// TIA Portal V21 export
// export: Created 2026-11-10T07:26:50.592199Z, ExportSetting WithDefaults, DisplayName Totally Integrated Automation Portal, DisplayVersion V21 Update 3, DisplayName STEP 7 Professional, DisplayVersion V21 Update 3, DisplayName STEP 7 Safety, DisplayVersion V21, DisplayName Tech WebApplication, DisplayVersion V21, DisplayName WinCC Basic/Comfort/Advanced, DisplayVersion V21 Update 3, DisplayName WinCC Unified, DisplayVersion V21 Update 3
FUNCTION_BLOCK "FB_LadOperands"   // FB5, LAD
{ S7_Optimized_Access := 'TRUE' }
VERSION : 0.1
// stored: AutoNumber true, IsIECCheckEnabled false, IsRetainMemResEnabled false, MemoryReserve 100, SetENOAutomatically false, UDAEnableTagReadback false
   VAR_INPUT
      "a" : Bool;
      ia : Int;
      wa : Word;
   END_VAR
   VAR_OUTPUT
      q : Bool;
      io : Int;
      dout : DInt;
      rout : Real;
      tout : Time;
      sout : String;
   END_VAR
   VAR_IN_OUT
      arr : Array[0..9] of Int;
   END_VAR
   VAR CONSTANT
      cInt : Int := 7;
   END_VAR
BEGIN

REGION Network 1: Absolute address word
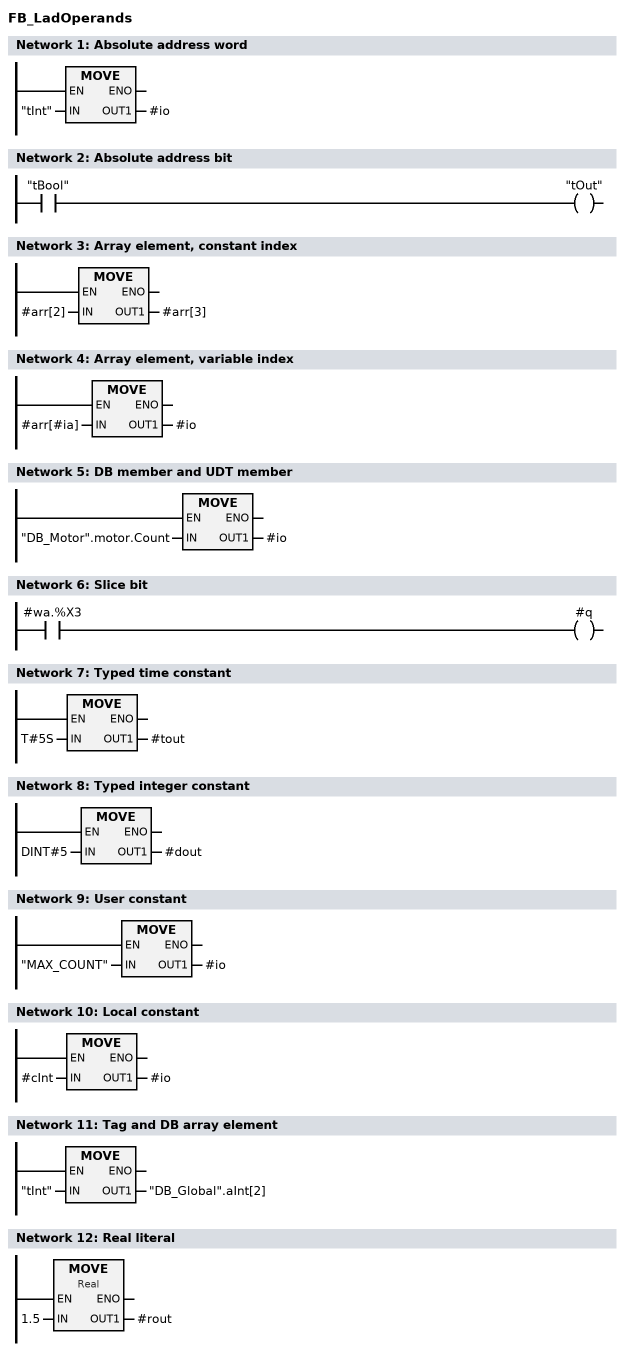
   RUNG wire#powerrail
      Move(in := "tInt", out1 => #io)
   END_RUNG
   // the same network as SCL:
   #io := "tInt";
END_REGION

REGION Network 2: Absolute address bit
   RUNG wire#powerrail
      Contact( "tBool" )
      Coil( "tOut" )
   END_RUNG
   // the same network as SCL:
   "tOut" := "tBool";
END_REGION

REGION Network 3: Array element, constant index
   RUNG wire#powerrail
      Move(in := #arr[2], out1 => #arr[3])
   END_RUNG
   // the same network as SCL:
   #arr[3] := #arr[2];
END_REGION

REGION Network 4: Array element, variable index
   RUNG wire#powerrail
      Move(in := #arr[#ia], out1 => #io)
   END_RUNG
   // the same network as SCL:
   #io := #arr[#ia];
END_REGION

REGION Network 5: DB member and UDT member
   RUNG wire#powerrail
      Move(in := "DB_Motor".motor.Count, out1 => #io)
   END_RUNG
   // the same network as SCL:
   #io := "DB_Motor".motor.Count;
END_REGION

REGION Network 6: Slice bit
   RUNG wire#powerrail
      Contact( #wa.%X3 )
      Coil( #q )
   END_RUNG
   // the same network as SCL:
   #q := #wa.%X3;
END_REGION

REGION Network 7: Typed time constant
   RUNG wire#powerrail
      Move(in := T#5S, out1 => #tout)
   END_RUNG
   // the same network as SCL:
   #tout := T#5S;
END_REGION

REGION Network 8: Typed integer constant
   RUNG wire#powerrail
      Move(in := DINT#5, out1 => #dout)
   END_RUNG
   // the same network as SCL:
   #dout := DINT#5;
END_REGION

REGION Network 9: User constant
   RUNG wire#powerrail
      Move(in := "MAX_COUNT", out1 => #io)
   END_RUNG
   // the same network as SCL:
   #io := "MAX_COUNT";
END_REGION

REGION Network 10: Local constant
   RUNG wire#powerrail
      Move(in := #cInt, out1 => #io)
   END_RUNG
   // the same network as SCL:
   #io := #cInt;
END_REGION

REGION Network 11: Tag and DB array element
   RUNG wire#powerrail
      Move(in := "tInt", out1 => "DB_Global".aInt[2])
   END_RUNG
   // the same network as SCL:
   "DB_Global".aInt[2] := "tInt";
END_REGION

REGION Network 12: Real literal
   RUNG wire#powerrail
      { S7_Templates := "SrcType := Real" } Move(in := 1.5, out1 => #rout)
   END_RUNG
   // the same network as SCL:
   #rout := 1.5;
END_REGION
END_FUNCTION_BLOCK
